(* IEC 61131-3 sources: JingjiangMoonbox/Application/Application/任务列表/Main_Task/IO配置表_1/QINHUA, 7 files *)

(* ---- KS_AbsEncModule_IODeal_QINHUA.st ---- *)
(*@CES
Name=KS_AbsEncModule_IODeal_QINHUA
Type=FunctionBlock
TypeGuid=6f9dac99-8de1-4efc-8465-68ac443b7d08
Guid=15f4a108-7592-45d5-8875-24926f1daf0a
HasDeclaration=True
HasImplementation=False
*)
{DECLARATION}
FUNCTION_BLOCK KS_AbsEncModule_IODeal_QINHUA
VAR_INPUT
	i_xInputEn:BOOL;
	i_xOutPutEn:BOOL;
	(*这些值的处理未考虑双收双放*)
	i_pdwAbsEncSinglePos_Uw:POINTER TO DWORD;
	i_pwAbsEncMultiPos_Uw:POINTER TO WORD;
	(*收料*)
	i_pdwAbsEncSinglePos_Rw:POINTER TO DWORD;
	i_pwAbsEncMultiPos_Rw:POINTER TO WORD;
	//2025.08.20.152113+
	i_pstStAbsEncIOModule_Uw:POINTER TO StAbsEncIOModule;
	i_pstStAbsEncIOModule_Rw:POINTER TO StAbsEncIOModule;

END_VAR
VAR
	wIWTest:WORD;
	wQWTest: WORD;
	byAbsEncSts: BOOL;
END_VAR

{IMPLEMENTATION}

(* ---- KS_FB_IOMAP_AIAO_QINHUA.st ---- *)
(*@CES
Name=KS_FB_IOMAP_AIAO_QINHUA
Type=FunctionBlock
TypeGuid=6f9dac99-8de1-4efc-8465-68ac443b7d08
Guid=95805f6d-5389-4683-9ccd-89bb7210177c
HasDeclaration=True
HasImplementation=False
*)
{DECLARATION}
FUNCTION_BLOCK KS_FB_IOMAP_AIAO_QINHUA
VAR_INPUT
	i_xEn: BOOL;(*功能块使能|*)
	i_xRdInput: BOOL;(*读io输入|*)
	i_xWrOutput: BOOL;(*写io输出|*)
	i_pstStSysParam								: POINTER TO StSysParam;
	i_pastStProgMonitoring						: POINTER TO ARRAY [1..2] OF StProgMonitoring;
END_VAR
VAR_OUTPUT
	o_xEno: BOOL;(*indicated to i_xEn|*)
	o_iErNo: INT;(*0.no err\-1.bad parameter|*)
END_VAR
VAR
//	fb_KS_FB_SetAIType: KS_FB_SetAIType;
	fbKS_FB_Analog_IO_CTL: KS_FB_Analog_IO_CTL;

	byAiFilterTms_UwRw_I					:  BYTE:= 1;(*滤波次数*)
	byAiFilterTms_UwRw_II					:  BYTE:= 1;
	byAiFilterTms_IfOf_I					:  BYTE:= 1;
	byAiFilterTms_IfOf_II					:  BYTE:= 1;
	byAiFilterTms_DiaMeasure_I				:   BYTE:= 1;
	byAiFilterTms_DiaMeasure_II				:   BYTE:= 1;
END_VAR

{IMPLEMENTATION}

(* ---- KS_FB_IOMAP_Axis_QINHUA.st ---- *)
(*@CES
Name=KS_FB_IOMAP_Axis_QINHUA
Type=FunctionBlock
TypeGuid=6f9dac99-8de1-4efc-8465-68ac443b7d08
Guid=0d2e69aa-ce38-4304-9029-5e42e440eb5b
HasDeclaration=True
HasImplementation=False
*)
{DECLARATION}
FUNCTION_BLOCK KS_FB_IOMAP_Axis_QINHUA
VAR_INPUT
	i_xEn: BOOL;(*功能块使能|*)
	i_xRdInput: BOOL;(*读io输入|*)
	i_xWrOutput: BOOL;(*写io输出|*)
	i_pastStIOMap_Axis_FE						: POINTER TO ARRAY [1..MAX_UNIT_NUM] OF StIOMap_Axis_FE;(*轴io数据区域|*)
END_VAR
VAR_OUTPUT
	o_xEno										: BOOL;(*indicated to i_xEn|*)
	o_iErNo										: INT;(*0.no err\-1.bad parameter|*)
END_VAR
VAR
	afbKS_FB_IOMap_Axis							: ARRAY [1..MAX_UNIT_NUM] OF KS_FB_MapAxisIOBasic;(*色组IO配置*)
END_VAR

{IMPLEMENTATION}

(* ---- KS_FB_IOMAP_AxisExtra_QINHUA.st ---- *)
(*@CES
Name=KS_FB_IOMAP_AxisExtra_QINHUA
Type=FunctionBlock
TypeGuid=6f9dac99-8de1-4efc-8465-68ac443b7d08
Guid=9bc3f83a-ed30-48fd-b56f-7d7783b3359f
HasDeclaration=True
HasImplementation=False
*)
{DECLARATION}
FUNCTION_BLOCK KS_FB_IOMAP_AxisExtra_QINHUA
VAR_INPUT
	i_xEn: BOOL;(*功能块使能|*)
	i_xRdInput: BOOL;(*读io输入|*)
	i_xWrOutput: BOOL;(*写io输出|*)
	i_pastStIOMap_Axis_Extra_FE						: POINTER TO ARRAY [1..MAX_UNIT_NUM] OF StIOMap_Axis_Extra_FE;(*轴io数据区域|*)
END_VAR
VAR_OUTPUT
	o_xEno										: BOOL;(*indicated to i_xEn|*)
	o_iErNo										: INT;(*0.no err\-1.bad parameter|*)
END_VAR
VAR
	afbKS_FB_IOMap_AxisExtra							: ARRAY [1..MAX_UNIT_NUM] OF KS_FB_MapAxisIOExtra;(*色组IO配置*)
END_VAR

{IMPLEMENTATION}

(* ---- KS_FB_IOMAP_Main_QINHUA.st ---- *)
(*@CES
Name=KS_FB_IOMAP_Main_QINHUA
Type=FunctionBlock
TypeGuid=6f9dac99-8de1-4efc-8465-68ac443b7d08
Guid=ef46cf9d-581d-4308-a97f-883e04346a23
HasDeclaration=True
HasImplementation=False
*)
{DECLARATION}
FUNCTION_BLOCK KS_FB_IOMAP_Main_QINHUA
(*主面板IO配置分A/B系和放/收牵*)
(*正常单收单放选1和2*)
(*双收双放1和2是A系的放牵收牵，3和4是B系的放牵收牵*)
(*双收双放A放B收1和4*)
VAR_INPUT
	i_xEn: BOOL;(*功能块使能|*)
	i_xRdInput: BOOL;(*读io输入|*)
	i_xWrOutput: BOOL;(*写io输出|*)
	i_pastStIOMap_Main_FE						: POINTER TO ARRAY [1..4] OF StIOMap_Main_FE;(*轴io数据区域|*)
END_VAR
VAR_OUTPUT
	o_xEno										: BOOL;(*indicated to i_xEn|*)
	o_iErNo										: INT;(*0.no err\-1.bad parameter|*)
END_VAR
VAR
	afbKS_FB_MapIO_Main						: ARRAY [1..4] OF KS_FB_MapIO_Main;(*主面板IO配置*)
END_VAR

{IMPLEMENTATION}

(* ---- KS_FB_IOMAP_UwRw_QINHUA.st ---- *)
(*@CES
Name=KS_FB_IOMAP_UwRw_QINHUA
Type=FunctionBlock
TypeGuid=6f9dac99-8de1-4efc-8465-68ac443b7d08
Guid=3e004c5e-d452-430c-a067-9e5d06a2c2c7
HasDeclaration=True
HasImplementation=False
*)
{DECLARATION}
 FUNCTION_BLOCK KS_FB_IOMAP_UwRw_QINHUA
VAR_INPUT
	i_xEn: BOOL;(*功能块使能|*)
	i_xRdInput: BOOL;(*读io输入|*)
	i_xWrOutput: BOOL;(*写io输出|*)
	i_pastStIOMap_UwRw_FE_Uw					: POINTER TO ARRAY [1..2] OF StIOMap_UwRw_FE;(*轴io数据区域|*)
	i_pastStIOMap_UwRw_FE_Rw					: POINTER TO ARRAY [1..2] OF StIOMap_UwRw_FE;(*轴io数据区域|*)
END_VAR
VAR_OUTPUT
	o_xEno										: BOOL;(*indicated to i_xEn|*)
	o_iErNo										: INT;(*0.no err\-1.bad parameter|*)
END_VAR
VAR
	afbKS_FB_MapIO_UwRw_Uw						: ARRAY [1..2] OF KS_FB_MapIO_UwRw;
	afbKS_FB_MapIO_UwRw_Rw						: ARRAY [1..2] OF KS_FB_MapIO_UwRw;
END_VAR

{IMPLEMENTATION}

(* ---- KS_FB_StepDriveIODeal_QINHUA.st ---- *)
(*@CES
Name=KS_FB_StepDriveIODeal_QINHUA
Type=FunctionBlock
TypeGuid=6f9dac99-8de1-4efc-8465-68ac443b7d08
Guid=93f5d248-e348-421d-8c6f-2346efeb17cc
HasDeclaration=True
HasImplementation=False
*)
{DECLARATION}
FUNCTION_BLOCK KS_FB_StepDriveIODeal_QINHUA
VAR_INPUT
	i_xInputEn:BOOL;
	i_xOutPutEn:BOOL;
	i_pastStDigitalMicroStepDrive :POINTER TO  ARRAY [1..MAX_UNIT_NUM] OF StDigitalMicroStepDrive;
	i_pastStStepDriveIOModule:POINTER TO ARRAY [1..MAX_UNIT_NUM] OF StStepDriveIOModule;
	i_pastStEnc0410R:POINTER TO ARRAY [1..MAX_UNIT_NUM] OF StEnc0410R;
END_VAR
VAR_OUTPUT
END_VAR
VAR
	wTest: WORD;
	afbKS_FB_StepDriveIOModule: ARRAY [1..MAX_UNIT_NUM] OF KS_FB_StepDriveIOModule;
END_VAR

{IMPLEMENTATION}
